{region 'Documentation'}
(*!
<summary>Checks whether text starts with the expected prefix, case-sensitively.</summary>
<description>

Read-only text must remain stable during the call and fit the configured Param_Assertions
text capacity. Invalid references or a missing terminator within that capacity report
Error.

The searched fragment, prefix or suffix must be nonempty; empty search text reports
Error. Matching is case-sensitive, without trimming or wildcard rules.

Diagnostic previews are shortened; the comparison still covers the complete validated
text.

</description>
*)
{endregion}
FUNCTION_BLOCK AssertStartsWith_String EXTENDS AssertionBase
VAR_IN_OUT CONSTANT
    IN : STRING(Param_Assertions.AssertionStringLength); //! Actual text.
    Prefix : STRING(Param_Assertions.AssertionStringLength); //! Expected prefix; must not be empty.
END_VAR

SUPER^();

{region 'Documentation'}
(*!
<summary>Validates inputs before comparing and escalating the result.</summary>
*)
{endregion}
METHOD PROTECTED Assert
VAR
    Message : STRING(GVL_Constants.MessageLength);
    PrefixText : STRING(GVL_Constants.AssertionValueLength);
    ActualText : STRING(GVL_Constants.AssertionValueLength);
END_VAR
IF NOT EvaluationActive THEN
    RETURN;
END_IF;

IF Result = E_Result.Error THEN
    RETURN;
END_IF;

// C0371: FB inputs are checked here before any reference access.
{warning disable C0371}
IF NOT __ISVALIDREF(IN) THEN
    Error(Message := 'Assertion error: IN reference is invalid.');
    RETURN;
END_IF;

IF NOT __ISVALIDREF(Prefix) THEN
    Error(Message := 'Assertion error: Prefix reference is invalid.');
    RETURN;
END_IF;

IF NOT IsAssertionStringLengthValid(Value := IN) THEN
    Error(Message := 'Assertion error: IN exceeds configured STRING length.');
    RETURN;
END_IF;

IF NOT IsAssertionStringLengthValid(Value := Prefix) THEN
    Error(Message := 'Assertion error: Prefix exceeds configured STRING length.');
    RETURN;
END_IF;

IF Prefix = '' THEN
    Error(Message := 'Assertion error: Prefix must not be empty.');
    RETURN;
END_IF;

IF Result = E_Result.Failed THEN
    RETURN;
END_IF;

IF NOT TextStartsWith_String(Value := IN,
    Prefix := Prefix) THEN
    PrefixText := CreateAssertionTextValue_String(Value := Prefix);
    ActualText := CreateAssertionTextValue_String(Value := IN);
    Message := CONCAT('Assertion failed: text does not start with expected prefix. Prefix = ',
        PrefixText);
    Message := CONCAT(Message, ', Actual = ');
    Message := CONCAT(Message, ActualText);
    Message := CONCAT(Message, '.');
    Fail(Message := Message);
    RETURN;
END_IF;

Pass();
{warning restore C0371}
END_METHOD

END_FUNCTION_BLOCK

(* stored: Version 1.1.0.1
   POU AssertStartsWith_String: Id {3994b2bb-80a3-4782-872b-fbc3d6f82019}, SpecialFunc None
   Folder Internal: Id {3cb07741-596b-46c7-b3e4-1bd91eb7b361}
   Method Assert: Id {9e4076e0-9f76-4788-a7e6-68a3864f1732} *)
